// TIA Portal V20 export
TYPE "Schrittkettensteuerung"
   STRUCT
      SK_Freigabe_Richten : Bool;
      SK_Richten_gestartet : Bool;
      SK_Richten_fertig : Bool;
      SK_Freigabe_Auto : Bool;
      SK_Aktiv : Bool;
      SK_Fertig : Bool;
      SK_Freigabe_Manuell_Auto : Bool;
      SK_Freigabe_Manuell_Richten : Bool;
      Reset_Freigaben : Bool;
      Station_1Ein_0Aus : Bool;
      SK_Richten_erforderlich : Bool;
      SK_Halt_von_Betriebsart : Bool;
   END_STRUCT;
END_TYPE
